// TIA Portal V20 export
DATA_BLOCK "HMI_SYS"   // DB2001
{ S7_Optimized_Access := 'FALSE' }
// stored: AutoNumber false
   VAR
      "Aktueller Bildschirm" : DInt := 1;
      Bildschirmwechsel : DInt := 1;
      Screen_Name : WString[254];
   END_VAR
BEGIN
END_DATA_BLOCK
